TEXTLIST TL_Test
  0 = 'Manual'
  1 = 'Semi-Auto'
  2 = 'Automatic'
   = ''
END_TEXTLIST

(* stored: Version 1.1.0.1
   TextList TL_Test: Id {68808e57-5b5b-468d-aecc-c52be0a9b605} *)
